// TIA Portal V20 export
Screen "190RB06_Stand_V23"  1276x673
  ScreenItem "Line_Header_X0_Y64" at 0,64 size 1276x0  Type=HmiLine
  ScreenItem "permanentareaborderrectangle" at 0,0 size 0x0  Type=HmiRectangle
  ScreenItem "Button_Back" at 2,2 size 90x60  Type=HmiButton
  ScreenItem "Title_ScreenOverview_X390_Y2_1" at 390,3 size 510x57  Type=HmiTextBox
  ScreenItem "Title_ScreenOverview_X390_Y2_5" at 1130,78 size 139x57  Type=HmiTextBox
  ScreenItem "Title_ScreenOverview_X390_Y2_6" at 1130,144 size 139x57  Type=HmiTextBox
  ScreenItem "Title_ScreenOverview_X390_Y2_7" at 1130,144 size 139x57  Type=HmiTextBox
  ScreenItem "Fusszeile_Button_ManualOPMode1_1" at 1088,2 size 90x60  Type=HmiButton
  ScreenItem "Fusszeile_Button_ManualOPMode1_4" at 1181,2 size 90x60  Type=HmiButton
  ScreenItem "Graphic view_1" at 457,157 size 358x495  Type=HmiGraphicView
  ScreenItem "Line_10" at 750,182 size 156x19  Type=HmiLine
  ScreenItem "Line_4" at 772,394 size 72x17  Type=HmiLine
  ScreenItem "Line_1" at 335,348 size 122x16  Type=HmiLine
  ScreenItem "文本域_11" at 201,308 size 134x40  Type=HmiTextBox
  ScreenItem "Rectangle_1" at 0,0 size 152x48  Type=HmiRectangle
  ScreenItem "文本域_1" at 2,1 size 122x45  Type=HmiTextBox
  ScreenItem "圆_1" at 0,0 size 100x30  Type=HmiCircle
  ScreenItem "圆_2" at 0,0 size 100x30  Type=HmiCircle
  ScreenItem "Rectangle_13" at 0,0 size 152x48  Type=HmiRectangle
  ScreenItem "文本域_19" at 2,1 size 122x45  Type=HmiTextBox
  ScreenItem "圆_5" at 0,0 size 100x30  Type=HmiCircle
  ScreenItem "圆_6" at 0,0 size 100x30  Type=HmiCircle
  ScreenItem "Title_ScreenOverview_X390_Y2_44" at 241,348 size 52x19  Type=HmiTextBox
  ScreenItem "Title_ScreenOverview_X390_Y2_46" at 268,368 size 25x21  Type=HmiTextBox
  ScreenItem "Title_ScreenOverview_X390_Y2_45" at 241,368 size 25x21  Type=HmiTextBox
